DATA_BLOCK "ControlNodes"
{ S7_Optimized_Access := 'TRUE' }
VERSION : 0.1
NON_RETAIN
STRUCT
    sequence : "LAF_typeSequence";
    jobs : "LAF_typeJobs";
    cylIZ02ExtPos : "LBC_TwoWayActuatorControlNodes";
    cylIZ02RetPos : "LBC_TwoWayActuatorControlNodes";
    cylQCamCoverExt : "LBC_TwoWayActuatorControlNodes";
    cylQCamCoverRet : "LBC_TwoWayActuatorControlNodes";
END_STRUCT;
BEGIN
END_DATA_BLOCK
